PROGRAM PRG_IntegrationScratch
VAR
END_VAR

; // integration-test scratch POU. Body is freely overwritten and restored by the live test suite. Never put real logic here.

END_PROGRAM

(* stored: Version 1.1.0.1
   POU PRG_IntegrationScratch: Id {2f32e079-63f9-4f56-9535-520b675581a8}, SpecialFunc None *)
